(* IEC 61131-3 sources: kns-port-domestic/targets/astra/lib/src/Interfaces/I_AlarmSink, 1 file *)

(* ---- OnAlarmEvent.method.decl.st ---- *)
// Событие перехода тревоги; FALSE — приёмник переполнен (FB_Alarm результат не повторяет)
METHOD OnAlarmEvent : BOOL
VAR_IN_OUT CONSTANT
    stEvent : ST_AlarmEvent;   // событие
END_VAR
